(* IEC 61131-3 sources: llm-plc-st-eval/data/processed_definitivo/claude-sonnet-4-6/C4/zero_shot, 3 files *)

(* ---- ejec_1.st ---- *)
FUNCTION_BLOCK FB_D

(* ─────────────────────────────────────────────────────────────────
   Entradas del bloque
   ───────────────────────────────────────────────────────────────── *)
VAR_INPUT
    demanda : BOOL;   (* Señal de demanda de bombeo (TRUE = se requiere caudal) *)
    falla1  : BOOL;   (* Señal de fallo de la Bomba 1 (TRUE = bomba en falla)   *)
    falla2  : BOOL;   (* Señal de fallo de la Bomba 2 (TRUE = bomba en falla)   *)
END_VAR

(* ─────────────────────────────────────────────────────────────────
   Salidas del bloque
   ───────────────────────────────────────────────────────────────── *)
VAR_OUTPUT
    bomba1   : BOOL;  (* Comando de arranque de la Bomba 1 (TRUE = arrancar)    *)
    bomba2   : BOOL;  (* Comando de arranque de la Bomba 2 (TRUE = arrancar)    *)
    almFalla : BOOL;  (* Alarma activa cuando la bomba prioritaria está en falla *)
END_VAR

(* ─────────────────────────────────────────────────────────────────
   Variables internas
   ───────────────────────────────────────────────────────────────── *)
VAR
    turno : BOOL;      (* Bit de turno: FALSE = prioridad Bomba 2,
                                        TRUE  = prioridad Bomba 1             *)
    fDem  : R_TRIG;    (* Detector de flanco ascendente sobre la señal demanda  *)
END_VAR

(* ─────────────────────────────────────────────────────────────────
   SECCIÓN 1 – Detección de flanco ascendente en la demanda
   Cada vez que 'demanda' pasa de FALSE a TRUE se genera un pulso
   en fDem.Q, lo que provoca la alternancia de turno.
   ───────────────────────────────────────────────────────────────── *)
fDem(CLK := demanda);

(* ─────────────────────────────────────────────────────────────────
   SECCIÓN 2 – Alternancia de turno
   Con cada nuevo flanco de demanda se invierte el bit 'turno',
   asegurando que las bombas se alternen como unidad prioritaria
   en cada ciclo de demanda consecutivo.
   ───────────────────────────────────────────────────────────────── *)
IF fDem.Q THEN
    turno := NOT turno;
END_IF

(* ─────────────────────────────────────────────────────────────────
   SECCIÓN 3 – Lógica de arranque y gestión de fallos
   ───────────────────────────────────────────────────────────────── *)
IF demanda THEN

    (* ── Rama A: turno = TRUE → Bomba 1 es la unidad prioritaria ── *)
    IF turno THEN
        (* Bomba 1 arranca si NO está en falla (es la prioritaria)   *)
        bomba1 := NOT falla1;

        (* Bomba 2 arranca como respaldo SOLO si Bomba 1 falló
           y Bomba 2 no tiene falla propia                           *)
        bomba2 := falla1 AND NOT falla2;

        (* Alarma activa si la unidad prioritaria (Bomba 1) falló    *)
        almFalla := falla1;

    (* ── Rama B: turno = FALSE → Bomba 2 es la unidad prioritaria ── *)
    ELSE
        (* Bomba 2 arranca si NO está en falla (es la prioritaria)   *)
        bomba2 := NOT falla2;

        (* Bomba 1 arranca como respaldo SOLO si Bomba 2 falló
           y Bomba 1 no tiene falla propia                           *)
        bomba1 := falla2 AND NOT falla1;

        (* Alarma activa si la unidad prioritaria (Bomba 2) falló    *)
        almFalla := falla2;
    END_IF

(* ─────────────────────────────────────────────────────────────────
   SECCIÓN 4 – Sin demanda: apagado total y reset de alarma
   Cuando no hay demanda ambas bombas se detienen y la alarma
   se desactiva, independientemente del estado de fallos.
   ───────────────────────────────────────────────────────────────── *)
ELSE
    bomba1   := FALSE;
    bomba2   := FALSE;
    almFalla := FALSE;
END_IF

END_FUNCTION_BLOCK

(* ---- ejec_2.st ---- *)
FUNCTION_BLOCK FB_D

(* ─────────────────────────────────────────────────────────────────────────
   Entradas del bloque
   ───────────────────────────────────────────────────────────────────────── *)
VAR_INPUT
    demanda : BOOL;   (* Señal de solicitud de bombeo (TRUE = hay demanda) *)
    falla1  : BOOL;   (* Señal de falla de la bomba 1 (TRUE = bomba 1 en falla) *)
    falla2  : BOOL;   (* Señal de falla de la bomba 2 (TRUE = bomba 2 en falla) *)
END_VAR

(* ─────────────────────────────────────────────────────────────────────────
   Salidas del bloque
   ───────────────────────────────────────────────────────────────────────── *)
VAR_OUTPUT
    bomba1   : BOOL;  (* Comando de arranque de la bomba 1 (TRUE = arrancar) *)
    bomba2   : BOOL;  (* Comando de arranque de la bomba 2 (TRUE = arrancar) *)
    almFalla : BOOL;  (* Alarma de falla activa en la bomba principal del turno *)
END_VAR

(* ─────────────────────────────────────────────────────────────────────────
   Variables internas
   ───────────────────────────────────────────────────────────────────────── *)
VAR
    turno : BOOL;    (* Indicador de turno: FALSE = bomba 2 es principal,
                                            TRUE  = bomba 1 es principal *)
    fDem  : R_TRIG;  (* Detector de flanco ascendente sobre la señal de demanda *)
END_VAR

(* ─────────────────────────────────────────────────────────────────────────
   SECCIÓN 1 – Detección de flanco ascendente en la señal de demanda
   Cada vez que 'demanda' pasa de FALSE a TRUE se genera un pulso en fDem.Q,
   lo que indica un nuevo ciclo de solicitud de bombeo.
   ───────────────────────────────────────────────────────────────────────── *)
fDem(CLK := demanda);

(* ─────────────────────────────────────────────────────────────────────────
   SECCIÓN 2 – Alternancia de turno
   En cada flanco ascendente de demanda se invierte 'turno', logrando que
   las bombas se alternen como unidad principal en cada nueva solicitud.
   ───────────────────────────────────────────────────────────────────────── *)
IF fDem.Q THEN
    turno := NOT turno;
END_IF

(* ─────────────────────────────────────────────────────────────────────────
   SECCIÓN 3 – Lógica de control de bombas según demanda y turno
   ───────────────────────────────────────────────────────────────────────── *)
IF demanda THEN

    (* ── Turno de bomba 1 como unidad principal ── *)
    IF turno THEN
        (* Bomba 1 arranca si NO tiene falla propia *)
        bomba1 := NOT falla1;

        (* Bomba 2 actúa como respaldo: arranca solo si bomba 1 falló
           Y bomba 2 no tiene falla propia *)
        bomba2 := falla1 AND NOT falla2;

        (* Alarma activa si la unidad principal (bomba 1) está en falla *)
        almFalla := falla1;

    (* ── Turno de bomba 2 como unidad principal ── *)
    ELSE
        (* Bomba 2 arranca si NO tiene falla propia *)
        bomba2 := NOT falla2;

        (* Bomba 1 actúa como respaldo: arranca solo si bomba 2 falló
           Y bomba 1 no tiene falla propia *)
        bomba1 := falla2 AND NOT falla1;

        (* Alarma activa si la unidad principal (bomba 2) está en falla *)
        almFalla := falla2;
    END_IF

(* ─────────────────────────────────────────────────────────────────────────
   SECCIÓN 4 – Sin demanda: apagado total y silencio de alarma
   ───────────────────────────────────────────────────────────────────────── *)
ELSE
    bomba1   := FALSE;  (* Detener bomba 1 *)
    bomba2   := FALSE;  (* Detener bomba 2 *)
    almFalla := FALSE;  (* Desactivar alarma *)
END_IF

END_FUNCTION_BLOCK

(* ---- ejec_3.st ---- *)
FUNCTION_BLOCK FB_D

(* ─────────────────────────────────────────────────────────────────────────
   Entradas del bloque
   ───────────────────────────────────────────────────────────────────────── *)
VAR_INPUT
    demanda : BOOL;   (* Señal de solicitud de bombeo (TRUE = hay demanda activa)  *)
    falla1  : BOOL;   (* Señal de falla de la bomba 1 (TRUE = bomba 1 en falla)    *)
    falla2  : BOOL;   (* Señal de falla de la bomba 2 (TRUE = bomba 2 en falla)    *)
END_VAR

(* ─────────────────────────────────────────────────────────────────────────
   Salidas del bloque
   ───────────────────────────────────────────────────────────────────────── *)
VAR_OUTPUT
    bomba1   : BOOL;  (* Comando de arranque para la bomba 1 (TRUE = arrancar)     *)
    bomba2   : BOOL;  (* Comando de arranque para la bomba 2 (TRUE = arrancar)     *)
    almFalla : BOOL;  (* Alarma de falla: TRUE cuando la bomba principal del turno
                         ha fallado y se ha activado (o intentado) el respaldo     *)
END_VAR

(* ─────────────────────────────────────────────────────────────────────────
   Variables internas
   ───────────────────────────────────────────────────────────────────────── *)
VAR
    turno : BOOL;    (* Bandera de turno: FALSE → bomba 2 es principal,
                                          TRUE  → bomba 1 es principal.
                        Persiste entre ciclos para mantener la alternancia.       *)
    fDem  : R_TRIG;  (* Detector de flanco ascendente sobre la señal de demanda;
                        se usa para cambiar el turno solo en cada nueva solicitud *)
END_VAR

(* ─────────────────────────────────────────────────────────────────────────
   SECCIÓN 1 – Detección de flanco ascendente en la demanda
   Cada vez que 'demanda' pasa de FALSE a TRUE se genera un pulso en fDem.Q,
   lo que dispara el cambio de turno (alternancia de bomba principal).
   ───────────────────────────────────────────────────────────────────────── *)
fDem(CLK := demanda);

(* ─────────────────────────────────────────────────────────────────────────
   SECCIÓN 2 – Alternancia de turno
   En el flanco ascendente de la demanda se invierte la bandera 'turno',
   seleccionando así la bomba principal para este nuevo ciclo de servicio.
   ───────────────────────────────────────────────────────────────────────── *)
IF fDem.Q THEN
    turno := NOT turno;   (* Invierte el turno: cambia la bomba principal *)
END_IF

(* ─────────────────────────────────────────────────────────────────────────
   SECCIÓN 3 – Lógica de control de bombas
   Solo se actúan las bombas mientras exista demanda activa.
   ───────────────────────────────────────────────────────────────────────── *)
IF demanda THEN

    (* ── Turno de bomba 1 como principal ─────────────────────────────────
       bomba1 arranca si NO tiene falla (es la principal y está sana).
       bomba2 arranca como respaldo SOLO si bomba1 falló y bomba2 está sana.
       almFalla se activa si la principal (bomba1) ha fallado.
       ─────────────────────────────────────────────────────────────────── *)
    IF turno THEN
        bomba1   := NOT falla1;              (* Principal: ON si no hay falla1          *)
        bomba2   := falla1 AND NOT falla2;   (* Respaldo:  ON solo si falla1 y no falla2*)
        almFalla := falla1;                  (* Alarma:    activa si la principal falló  *)

    (* ── Turno de bomba 2 como principal ─────────────────────────────────
       bomba2 arranca si NO tiene falla (es la principal y está sana).
       bomba1 arranca como respaldo SOLO si bomba2 falló y bomba1 está sana.
       almFalla se activa si la principal (bomba2) ha fallado.
       ─────────────────────────────────────────────────────────────────── *)
    ELSE
        bomba2   := NOT falla2;              (* Principal: ON si no hay falla2          *)
        bomba1   := falla2 AND NOT falla1;   (* Respaldo:  ON solo si falla2 y no falla1*)
        almFalla := falla2;                  (* Alarma:    activa si la principal falló  *)
    END_IF

(* ─────────────────────────────────────────────────────────────────────────
   SECCIÓN 4 – Sin demanda
   Cuando no hay solicitud de bombeo se apagan ambas bombas y se silencia
   la alarma de falla, dejando el sistema en reposo seguro.
   ───────────────────────────────────────────────────────────────────────── *)
ELSE
    bomba1   := FALSE;   (* Apagar bomba 1 *)
    bomba2   := FALSE;   (* Apagar bomba 2 *)
    almFalla := FALSE;   (* Silenciar alarma *)
END_IF

END_FUNCTION_BLOCK
